TYPE "TiaMcpDepInner"
VERSION : 0.1
STRUCT
    Value : Int;
END_STRUCT;
END_TYPE
